PROGRAM MAIN
VAR
    Machine  : DemoMachine;
    Listener : AlarmListener;
END_VAR

Machine.CyclicLogic(Commands := GVL_Hmi.Commands, Status := GVL_Hmi.Status);
Listener.CyclicLogic(Table := GVL_Hmi.PlcAlarms);

END_PROGRAM

(* stored: Version 1.1.0.1, ProductVersion 3.1.4024.12
   POU MAIN: Id {95e5a0e8-cb77-4cfa-8792-3bcb5a7fec1a}, SpecialFunc None *)
